Staubli VAL3: onStart.pgx

public program onStart()
  local num l_i
begin
  call saveData:setBaseJOG(saveData:nJogTool)
  resize(sList,1,size(safeTemp:sSPoint))
  for l_i = 0 to size(sList)-1
    sList[l_i]=toString("",l_i)+","+safeTemp:sSPoint[l_i].sName
  endFor

  sSelPoint=""
  sLastPoint=""
  bActive=false

  for l_i = 0 to size(sTRSF)-1
    sTRSF[l_i]=""
  endFor

end
